(* IEC 61131-3 sources: SortJet_MasterSPS_Aufbau.fbsproj/09_Station/Stationen/_Allgemein, 5 files *)

(* ---- Arretierung_FB_V01_00_00.fb.st ---- *)
(* METADATA
{
	"v3Meta": {
		"objectGuid": "dcab1ddf-6c10-4772-a9bc-4c92780e70eb"
	}
}
*)
FUNCTION_BLOCK Arretierung_FB_V01_00_00
VAR_INPUT

  // EINGAENGE
  in_bStatusZylinderAusgefahren : BOOL;
  in_bStatusZylinderEingefahren : BOOL;

  // BOOLEAN
  bpReset                       : BOOL;
  bpAktivieren                  : BOOL;
  bpFreigabe                    : BOOL; // FREIGABE Pneumatik: ohne Freigabe Ventile aus, Bewegung pausiert (Startbefehl bleibt erhalten)
  bpStartAusfahren              : BOOL;
  bpStartEinfahren              : BOOL;

  // OPTIONEN
  bpAbfrageAusgefahrenVorhanden : BOOL := TRUE;   // Endlagensensor ausgefahren vorhanden, sonst gilt die Endlage nach tpBewegungszeit
  bpAbfrageEingefahrenVorhanden : BOOL := TRUE;   // Endlagensensor eingefahren vorhanden, sonst gilt die Endlage nach tpBewegungszeit
  tpBewegungszeit               : TIME := T#800MS; // Bewegungszeit je Richtung ohne Endlagensensor

END_VAR
VAR_OUTPUT
  // AUSGAENGE
  out_bZylinderAusfahren        : BOOL;
  out_bZylinderEinfahren        : BOOL;

  // BOOLEAN
  bpFehler                      : BOOL;
  bpDone                        : BOOL;

  // WORD
  wpFehlerNr                    : Fehlerkonstanten_EN;

  // ENUM
  epStatusZylinder : PneumatikZylinderStatus_EN;

END_VAR
VAR

  // STEPS
  steplAusfahren   : Steps_TE;
  steplEinfahren   : Steps_TE;

  // TIMER
  tonZylinderEingefahren     : TON; // EINSCHALTVERZOEGERUNG: Warten bis der Zylinder eingefahren wurde. Sonst wird ein Fehlerausgegeben
  tonZylinderAusgefahren     : TON; // EINSCHALTVERZOEGERUNG: Warten bis der Zylinder ausgefahren wurde. Sonst wird ein Fehlerausgegeben
  tonlBewegungszeitEinfahren : TON; // Bewegungszeit ohne Endlagensensor eingefahren
  tonlBewegungszeitAusfahren : TON; // Bewegungszeit ohne Endlagensensor ausgefahren

END_VAR

VAR CONSTANT

  // TIME
  cZEITLICHE_UEBERWACHUNG_BEWEGUNG_ZYLINDER : TIME := T#15s;

END_VAR
//-------------------------------------------------------------------------------------------------
// BAUSTEIN: RESET / DEAKTIVIERT
//-------------------------------------------------------------------------------------------------
(* Hinweis:
   - Reset oder deaktiviert: Ausgaenge aus, Ketten und Timer zuruecksetzen, Done und Fehler loeschen
   - Der Baustein setzt bpReset selbst zurueck, der Aufrufer wartet nicht auf Done
   - Ein deaktivierter Zylinder meldet kein Done; der Aufrufer verknuepft das Warten auf Done
     mit der Aktivierung aus der MK (z.B. Zylinder.bpDone OR NOT stStationsAufbau.bX)
*)
IF ( bpReset OR NOT bpAktivieren ) THEN

  out_bZylinderAusfahren := FALSE;
  out_bZylinderEinfahren := FALSE;

  bpStartAusfahren := FALSE;
  bpStartEinfahren := FALSE;

  steplAusfahren := STEP_0_E;
  steplEinfahren := STEP_0_E;

  tonZylinderAusgefahren( IN := FALSE );
  tonZylinderEingefahren( IN := FALSE );
  tonlBewegungszeitAusfahren( IN := FALSE );
  tonlBewegungszeitEinfahren( IN := FALSE );

  bpDone     := FALSE;
  bpFehler   := FALSE;
  wpFehlerNr := cMELDUNG_NULL;

  bpReset := FALSE;

  RETURN;

END_IF

//-------------------------------------------------------------------------------------------------
// BAUSTEIN: AKTIONEN
//-------------------------------------------------------------------------------------------------
(* Hinweis Freigabe Pneumatik:
   - Ohne Freigabe: Ventile aus, Ketten und Ueberwachungszeiten zuruecksetzen (kein Timeout-Fehler)
   - Der Startbefehl bleibt erhalten: kommt die Freigabe zurueck, wird die Bewegung neu gestartet
*)
IF NOT bpFreigabe THEN
  out_bZylinderAusfahren := FALSE;
  out_bZylinderEinfahren := FALSE;
  steplAusfahren := STEP_0_E;
  steplEinfahren := STEP_0_E;
  tonZylinderAusgefahren( IN := FALSE );
  tonZylinderEingefahren( IN := FALSE );
  tonlBewegungszeitAusfahren( IN := FALSE );
  tonlBewegungszeitEinfahren( IN := FALSE );
  bpDone := FALSE;
ELSE
  Ausfahren();
  Einfahren();
END_IF

//-------------------------------------------------------------------------------------------------
// STATUS DES ZYLINDERS
//-------------------------------------------------------------------------------------------------
(* Hinweis:
   - Status aus der Sensorik, soweit Endlagensensoren vorhanden sind
   - Ohne Sensor bleibt der Status, den die Schrittketten nach der Bewegungszeit setzen
*)
IF ( bpAbfrageAusgefahrenVorhanden AND bpAbfrageEingefahrenVorhanden ) THEN

  IF (      in_bStatusZylinderAusgefahren
       AND NOT in_bStatusZylinderEingefahren )
  THEN
    epStatusZylinder := eZylinderAusgefahren;
  ELSIF(    in_bStatusZylinderEingefahren
         AND NOT in_bStatusZylinderAusgefahren )
  THEN
    epStatusZylinder := eZylinderEingefahren;
  ELSE
    epStatusZylinder := eZylinderUndefiniert;
  END_IF

ELSIF ( bpAbfrageAusgefahrenVorhanden ) THEN

  IF ( in_bStatusZylinderAusgefahren ) THEN
    epStatusZylinder := eZylinderAusgefahren;
  ELSIF ( epStatusZylinder = eZylinderAusgefahren ) THEN
    epStatusZylinder := eZylinderUndefiniert;
  END_IF

ELSIF ( bpAbfrageEingefahrenVorhanden ) THEN

  IF ( in_bStatusZylinderEingefahren ) THEN
    epStatusZylinder := eZylinderEingefahren;
  ELSIF ( epStatusZylinder = eZylinderEingefahren ) THEN
    epStatusZylinder := eZylinderUndefiniert;
  END_IF

END_IF
END_FUNCTION_BLOCK

(* ---- Kippen_FB_V01_00_00.fb.st ---- *)
(* METADATA
{
	"v3Meta": {
		"objectGuid": "d572774f-9eb0-4642-b999-1d4bc3469776"
	}
}
*)
FUNCTION_BLOCK Kippen_FB_V01_00_00
VAR_INPUT

  // BOOLEAN *)
  bpAktivieren              : BOOL;
  bpFreigabe                : BOOL;
  bpReset                   : BOOL;
  bpReferenz                : BOOL;
  bpPositionieren           : BOOL;
  bpHandfahrenPlus          : BOOL;
  bpHandfahrenMinus         : BOOL;
  bpAutomatikAktiv          : BOOL;
  bpSensorEinlauf           : BOOL;
  bpSensorAuslauf           : BOOL;
  bpSensorEinlaufNachfolger : BOOL;
  bpSensorAuslaufVorgaenger : BOOL;
  bpTeilnehmerErreichbar    : BOOL;

  bpSensorNicht90Grad       : BOOL;

  bpLangsamKippen           : BOOL; // Umrichter: mit reduzierter Geschwindigkeit und Beschleunigung positionieren
  bpSensorNicht84Grad       : BOOL;

  // POINTER
  ppAntriebsInformationen : REFERENCE TO AntriebsInformationen;
  ppParameterBaustein     : REFERENCE TO Parameter_Kippen;

  // ENUM
  epZielPosition          : Kippen_EN; // Hinweis: Wird fuer die Absolut-Positionierung verwendet "bpStartAbsolutPositionierung"

  // STRUCT
  stStationsNummern       : Station_ST;

END_VAR
VAR_OUTPUT

  // BOOLEAN
  bpDone                       : BOOL;
  bpFehler                     : BOOL;
  bpInReferenz                 : BOOL;
  bpPositionierenAbgeschlossen : BOOL;

  // WORD
  wpFehlerNr                   : Fehlerkonstanten_EN; // FEHLER-AUSWERTUNG: Fehlernummer[Const] *)

  // ENUM *)
  epKippStatus                 : Kippen_EN; // Status: Gibt die aktuelle Position des Antriebs aus

END_VAR
VAR

  // BOOLEAN
  blErsterZyklus      : BOOL := TRUE;

  // REAL
  rlAntriebsZielPosition : REAL;

  // TIMER
  tonlFehlermeldungUnterdrueckenAntriebOK : TON;
  tonlMaxWarteZeit                        : TON;
  tonlMaxWarteAufResetErfolgreich         : TON;
  tonlAntriebNichtFreigegeben             : TON; // Ueberwachung: Antrieb nicht betriebsbereit
  tonlEndschalterFreifahren               : TON;
  tonlWarteSchrittEndschalterFreifahren   : TON;
  tofHardwareEndschalterFrei              : TOF;
  toflReglerFreigabeErhalten              : TOF;
  toflHardwareEndschalterFrei             : TOF;
  toflReset                               : TOF;

  // STEPS
  steplReset          : Steps_TE;
  steplReferenz       : Steps_TE;
  steplPositionieren  : Steps_TE;

  // Antrieb
  Antrieb : REFERENCE TO Rexroth_ctrlX_Drive_Eckelmann_MC_V01_02_02;

END_VAR

VAR
  // HARDWARE EINGÄNGE
  in_bMotorstarter_OK                 AT%I* : BOOL;
  in_bLS400V_OK                       AT%I* : BOOL;
  in_bLSBremse_OK                     AT%I* : BOOL;

  // HARDWARE AUSGÄNGE
  out_bKippen84Grad                   AT%Q* : BOOL;
  out_bKippen90Grad                   AT%Q* : BOOL;
  out_bBremseLoesen                   AT%Q* : BOOL;
  out_bReset                          AT%Q* : BOOL;

END_VAR

//-------------------------------------------------------------------------------------------------
// INITIALISIERUNG
//-------------------------------------------------------------------------------------------------
IF ( blErsterZyklus ) THEN

  IF ( __ISVALIDREF(ppAntriebsInformationen) ) THEN

    blErsterZyklus := FALSE;

    Antrieb REF= pgAntriebe[ppAntriebsInformationen.wAchsID];

    (* Hinweis:
       - Initialisierung Antriebsinformationen
    *)
    Antrieb.ppAntriebsInformationen REF= ppAntriebsInformationen;

    (* Hinweis:
       - Für die Zielpunktkontrolle muss im ersten Zyklus die Zielposition initialisiert werden
    *)
    Antrieb.rpZielPosition := Antrieb.rpIstPosition;

    (* Hinweis:
       - Antriebswerte vorinitialisieren
    *)
    Antrieb.rpGeschwindigkeit := ppAntriebsInformationen.rpMaxGeschwindigkeit;
    Antrieb.rpBeschleunigung  := ppAntriebsInformationen.rpMaxBeschleunigung;
    Antrieb.rpVerzoegerung    := ppAntriebsInformationen.rpMaxVerzoegerung;
    Antrieb.rpRuckzeit        := ppAntriebsInformationen.rpMaxRuckzeit;

  ELSE
    RETURN;
  END_IF

END_IF

//-------------------------------------------------------------------------------------------------
// DEAKTIVIEREN
//-------------------------------------------------------------------------------------------------
IF ( NOT bpAktivieren ) THEN

  bpDone                       := TRUE;
  bpInReferenz                 := TRUE;
  bpPositionierenAbgeschlossen := TRUE;

  epKippStatus := epZielPosition;

  bpFehler   := FALSE;
  wpFehlerNr := cMELDUNG_NULL;

  RETURN;

END_IF

//-------------------------------------------------------------------------------------------------
// BAUSTEIN: AKTIONEN
//-------------------------------------------------------------------------------------------------

(* Hinweis:
   - Kippbewegung
*)
IF (ppParameterBaustein.bKippenMitSchuetz ) THEN
  Kippen_Schuetz();
ELSE
  Positionieren();
END_IF

(* Hinweis:
   - Baisis- Aktionen
*)
Ausgaenge();
Meldungen();
Timer();
Reset();
Referenz();
Handbetrieb();

//-------------------------------------------------------------------------------------------------
// ZUWEISUNGEN UND BAUSTEINAUFRUFE
//-------------------------------------------------------------------------------------------------
// Antriebsfreigabe:
//    - Antrieb
toflReglerFreigabeErhalten( IN := (   bpPositionieren
                                    OR bpReferenz
                                    OR bpHandfahrenPlus
                                    OR bpHandfahrenMinus
                                    OR bpReset ),
                            PT := ppParameterBaustein.tZeitAntriebsfreigabeErhalten );

Antrieb.bpFreigabe        := ( bpFreigabe AND toflReglerFreigabeErhalten.Q );
IF ( NOT ( bpPositionieren AND bpLangsamKippen ) ) THEN
  Antrieb.rpRuckzeit      := ppAntriebsInformationen.rpMaxRuckzeit;
END_IF
Antrieb.stStationsNummern := stStationsNummern;
END_FUNCTION_BLOCK

(* ---- Messachse_FB_V01_00_00.fb.st ---- *)
(* METADATA
{
	"v3Meta": {
		"objectGuid": "ee8fce2f-1a3c-411c-afad-25d0a39b52dd"
	}
}
*)
FUNCTION_BLOCK Messachse_FB_V01_00_00
VAR_INPUT

  // BOOL
  bpAktivieren                             : BOOL;
  bpPositionierung                         : BOOL;
  bpVermessen_OberUndUnterkante_2_Sensoren : BOOL;
  bpVermessen_Oberkante_1_Sensor           : BOOL;
  bpReset                                  : BOOL;
  bpReferenz                               : BOOL;
  bpFreigabe                               : BOOL;
  bpHandfahrenPlus                         : BOOL;
  bpHandfahrenMinus                        : BOOL;
  bpBetriebsartHand                        : BOOL;
  bpFusstaster                             : BOOL;

 // REAL
  rpZielPosition                           : REAL;
  rpErwarteteScheibenHoehe                 : REAL;

  // STRUCT
  stStationsNummern                        : Station_ST;

  // POINTER
  ppAntriebsInformationen                  : REFERENCE TO AntriebsInformationen;
  ppParameterBaustein                      : REFERENCE TO Parameter_Messachse;

END_VAR
VAR_OUTPUT

  // BOOL
  bpDone                    : BOOL;
  bpFehler                  : BOOL;
  bpInReferenz              : BOOL;
  bprtScheibe               : BOOL;
  bpVermessenAbgeschlossen  : Bool;

  // WORD
  wpFehlerNr                : Fehlerkonstanten_EN;

  // REAL
  rpIstPosition             : REAL;
  rlScheibenunterkante      : REAL;
  rlScheibenoberkante       : REAL;
  rlMessErgebnis            : REAL;
  rlPositionAntriebBeiStart : REAL;
  rlBremsWeg                : REAL;

  // ENUM
  epGlashoehenTyp      : GlasHoehenTyp_EN;
  epGlashoehenTypMode2 : GlasHoehenTyp_EN;

END_VAR
VAR

  // BOOL
  blErsterZyklus                         : BOOL := TRUE;

  // REAL
  rlBremsPos                             : REAL;
  rlOffsetMinimumFrueherBremsen          : REAL := 150;
  rlOffsetMaximumFrueherBremsen          : REAL := 300;

  // TIMER
  tonlEndschalterFreifahren              : TON;
  tonlWarteSchrittEndschalterFreifahren  : TON;
  tonlMaxWarteAufResetErfolgreich        : TON;
  tonlAntriebNichtFreigegeben            : TON; // Ueberwachung: Antrieb nicht betriebsbereit
  tonlTimeoutUnterkante                  : TON;
  toflHardwareEndschalterFrei            : TOF;
  toflReglerFreigabeErhalten             : TOF;

  // STEPS
  steplPositionieren                     : Steps_TE;
  steplReferenz                          : Steps_TE;
  steplReset                             : Steps_TE;
  steplOberkante_1_Sensor                : Steps_TE;
  steplOberUndUnterkante_2_Sensoren      : Steps_TE;

  // Antrieb
  Antrieb : REFERENCE TO Rexroth_ctrlX_Drive_Eckelmann_MC_V01_02_02;

END_VAR

VAR_INPUT

  // HARDWARE EINGAENGE
  in_bSensorUnten                        : BOOL;
  in_bSensorOben                         : BOOL;
  in_bSensorUnterkante                   : BOOL;
  in_bEndschalterMin                     : BOOL; // Oeffner (TRUE = frei), gemappt; zum Umrichter ueber Signal-Steuerwort Bit 10, wirkt nur bei Endschalterquelle SPS

END_VAR
VAR CONSTANT

  // REAL
  cUEBERWACHUNG_WEGSTRECKE  : REAL := 40.0;

END_VAR

//-------------------------------------------------------------------------------------------------
// INITIALISIERUNG
//-------------------------------------------------------------------------------------------------
IF ( blErsterZyklus ) THEN

  IF ( __ISVALIDREF(ppAntriebsInformationen) ) THEN

    blErsterZyklus := FALSE;

    Antrieb REF= pgAntriebe[ppAntriebsInformationen.wAchsID];

    (* Hinweis:
       - Initialisierung Antriebsinformationen
    *)
    Antrieb.ppAntriebsInformationen REF= ppAntriebsInformationen;

    (* Hinweis:
       - Für die Zielpunktkontrolle muss im ersten Zyklus die Zielposition initialisiert werden
    *)
    Antrieb.rpZielPosition := Antrieb.rpIstPosition;

    (* Hinweis:
       - Antriebswerte vorinitialisieren
    *)
    Antrieb.rpGeschwindigkeit := ppAntriebsInformationen.rpMaxGeschwindigkeit;
    Antrieb.rpBeschleunigung  := ppAntriebsInformationen.rpMaxBeschleunigung;
    Antrieb.rpVerzoegerung    := ppAntriebsInformationen.rpMaxVerzoegerung;
    Antrieb.rpRuckzeit        := ppAntriebsInformationen.rpMaxRuckzeit;

  ELSE
    RETURN;
  END_IF

END_IF

//-------------------------------------------------------------------------------------------------
// DEAKTIVIEREN
//-------------------------------------------------------------------------------------------------
IF ( NOT bpAktivieren ) THEN

  bpDone := TRUE;

  (* Hinweis:
     - Ausnahmesituationen
  *)
  bpInReferenz := TRUE;
  bpFehler   := FALSE;
  wpFehlerNr := cMELDUNG_NULL;

  RETURN;

END_IF

//-------------------------------------------------------------------------------------------------
// IO's
//-------------------------------------------------------------------------------------------------
in_bSensorOben       := Antrieb.udipEingaengeUmrichter.cXG31_2_I_2;
in_bSensorUnten      := Antrieb.udipEingaengeUmrichter.cXG31_1_I_1;
in_bSensorUnterkante := Antrieb.udipEingaengeUmrichter.cXG37_4_I_6;
Antrieb.bpEndschalterMinExtern := in_bEndschalterMin;

//-------------------------------------------------------------------------------------------------
// BAUSTEIN: AKTIONEN
//-------------------------------------------------------------------------------------------------

Positionieren();
Vermessen_Oberkante_1_Sensor();
Vermessen_OberUndUnterkante_2_Sensoren();
Reset();
Referenz();
Handfunktion();

//-------------------------------------------------------------------------------------------------
// BAUSTEIN: AUSGAENGE
//-------------------------------------------------------------------------------------------------
// Ausgabe der Aktuellen Position
rpIstPosition := Antrieb.rpIstPosition;
bpInReferenz := Antrieb.bpIstReferenziert;

(* Hinweis:
   - Scheibenhoehe kontrollieren
*)
IF ( in_bSensorUnten AND NOT in_bSensorOben ) THEN
  epGlashoehenTyp := eGlasHoeheOK;

ELSE

  IF ( NOT in_bSensorUnten AND NOT in_bSensorOben ) THEN
    epGlashoehenTyp := eGlasZuNiedrig;

  ELSIF ( in_bSensorUnten AND  in_bSensorOben ) THEN
    epGlashoehenTyp := eGlasZuHoch;

  END_IF

END_IF

//-------------------------------------------------------------------------------------------------
// BAUSTEIN: AUFRUFE
//-------------------------------------------------------------------------------------------------
toflReglerFreigabeErhalten( IN := (   bpPositionierung
                                    OR bpReferenz
                                    OR bpHandfahrenPlus
                                    OR bpHandfahrenMinus
                                    OR bpVermessen_OberUndUnterkante_2_Sensoren
                                    OR bpVermessen_Oberkante_1_Sensor
                                    OR bpReset ),
                            PT := tgZeitAutoabschaltungEnergiesparModus );

Antrieb.bpFreigabe        := ( bpFreigabe AND toflReglerFreigabeErhalten.Q );
Antrieb.rpRuckzeit        := ppAntriebsInformationen.rpMaxRuckzeit;
Antrieb.stStationsNummern := stStationsNummern;

//-------------------------------------------------------------------------------------------------
// BAUSTEIN: AUSNAHMESITUATIONEN
//-------------------------------------------------------------------------------------------------
IF ( Antrieb.bpFehler
     AND NOT ( steplPositionieren = STEP_900_E
               OR steplOberUndUnterkante_2_Sensoren = STEP_900_E
               OR steplOberkante_1_Sensor = STEP_900_E
               OR steplReferenz    = STEP_900_E
               OR steplReset       = STEP_900_E ) )
THEN
  wpFehlerNR := cMELDUNG_ANTRIEB_MESSACHSE;
  bpFehler := TRUE;
END_IF
END_FUNCTION_BLOCK

(* ---- Querfahrt_FB_V01_00_00.fb.st ---- *)
(* METADATA
{
	"v3Meta": {
		"objectGuid": "62b3e7d5-59d7-4fa9-a26b-9f6c0e862cd9"
	}
}
*)
FUNCTION_BLOCK Querfahrt_FB_V01_00_00
VAR_INPUT

  // BOOLEAN
  bpAktivieren                           : BOOL;
  bpFreigabe                             : BOOL;
  bpAutomatikAktiv                       : BOOL;
  bpPositionieren                        : BOOL;
  bpReset                                : BOOL;
  bpReferenz                             : BOOL;
  bpHandfahrenPlus                       : BOOL;
  bpHandfahrenMinus                      : BOOL;

  bpSensorEinlauf                        : BOOL;
  bpSensorAuslauf                        : BOOL;
  bpSensorAuslaufVorgaenger              : BOOL;
  bpVerfahrfreigabe                      : BOOL := TRUE; // Externe Freigabe zum Verfahren (ohne Beschaltung TRUE)
  bpQuittungAuftragsstatusZurueckgesetzt : BOOL; // Auftrag wurde zurueckgesetzt
  bpReglungAktivSchalten                 : BOOL; // Da der Querfahrtantrieb keine Bremse hat, muss um die Position zu halten der Regler in Regelung stehen, sonst verschiebt sich die Station *)

  // REAL
  rpZielPosition                         : REAL;

  // POINTER
  ppParameterBaustein                    : REFERENCE TO Parameter_Querfahrt;
  ppAntriebsInformationen                : REFERENCE TO AntriebsInformationen;

  // STRUKTUR
  stStationsNummern                      : Station_ST;

END_VAR
VAR_OUTPUT

  // BOOLEAN
  bpDone                                 : BOOL;
  bpFehler                               : BOOL;
  bpAntrieblaeuft                        : BOOL;
  bpAuftragAktiv                         : BOOL;
  bpAuftragsstatusZuruecksetzen          : BOOL := FALSE;
  bpPositionierungGestartet              : BOOL := FALSE;
  bpPositionierungAbgeschlossen          : BOOL := FALSE;
  bpMinEndschalterBelegt                 : BOOL := FALSE;
  bpMaxEndschalterBelegt                 : BOOL := FALSE;
  bpZielPositionErreicht                 : BOOL;
  bpInReferenz                           : BOOL;

  // WORD
  wpFehlerNr                             : Fehlerkonstanten_EN;

  // REAL
  rpAktuellePosition                     : REAL;

END_VAR
VAR

  // BOOL
  blErsterZyklus                         : BOOL := TRUE;
  blVerfahrfreigabe                      : BOOL;
  blAbbruchPositionierung                : BOOL := FALSE;

  // STEPS
  steplPositionieren                     : Steps_TE;
  steplReferenz                          : Steps_TE;
  steplReset                             : Steps_TE;

  // TIMER
  tonlEndschalterFreifahren              : TON;
  tonlMaxWarteAufResetErfolgreich        : TON;
  toflHardwareEndschalterFrei            : TOF;
  toflReglerFreigabeErhalten             : TOF;

  // Antrieb
  Antrieb : REFERENCE TO Rexroth_ctrlX_Drive_Eckelmann_MC_V01_02_02;

END_VAR

//-------------------------------------------------------------------------------------------------
// INITIALISIERUNG
//-------------------------------------------------------------------------------------------------
IF ( blErsterZyklus ) THEN

  IF ( __ISVALIDREF(ppAntriebsInformationen) ) THEN

    blErsterZyklus := FALSE;

    Antrieb REF= pgAntriebe[ppAntriebsInformationen.wAchsID];

    (* Hinweis:
       - Initialisierung Antriebsinformationen
    *)
    Antrieb.ppAntriebsInformationen REF= ppAntriebsInformationen;

    (* Hinweis:
       - Für die Zielpunktkontrolle muss im ersten Zyklus die Zielposition initialisiert werden
    *)
    Antrieb.rpZielPosition := Antrieb.rpIstPosition;

    (* Hinweis:
       - Antriebswerte vorinitialisieren
    *)
    Antrieb.rpGeschwindigkeit := ppAntriebsInformationen.rpMaxGeschwindigkeit;
    Antrieb.rpBeschleunigung  := ppAntriebsInformationen.rpMaxBeschleunigung;
    Antrieb.rpVerzoegerung    := ppAntriebsInformationen.rpMaxVerzoegerung;
    Antrieb.rpRuckzeit        := ppAntriebsInformationen.rpMaxRuckzeit;

  ELSE
    RETURN;
  END_IF

END_IF

//-------------------------------------------------------------------------------------------------
// DEAKTIVIEREN
//-------------------------------------------------------------------------------------------------
IF ( NOT bpAktivieren ) THEN

  bpDone                        := TRUE;
  bpAuftragsstatusZuruecksetzen := FALSE;

  bpFehler   := FALSE;
  wpFehlerNr := cMELDUNG_NULL;

  RETURN;

END_IF

//-------------------------------------------------------------------------------------------------
// AKTIONEN
//-------------------------------------------------------------------------------------------------
// Verfahrfreigabe (lokal, der Eingang wird nicht ueberschrieben)
blVerfahrfreigabe :=     bpVerfahrfreigabe
                         AND NOT bpSensorEinlauf
                         AND NOT bpSensorAuslauf
                         AND NOT bpSensorAuslaufVorgaenger;

Verfahrlogik();
Positionieren();
Handfunktionen();
Reset();
Referenz();
Meldungen();

//-------------------------------------------------------------------------------------------------
// Freigabe zum Verfahren
//-------------------------------------------------------------------------------------------------
IF NOT blVerfahrfreigabe AND Antrieb.wpBetriebsart <> AntriebsBetriebsart_EN.RESET AND Antrieb.wpBetriebsart <> KEINE_FUNKTION THEN
  Antrieb.wpBetriebsart := KEINE_FUNKTION;
END_IF

//-------------------------------------------------------------------------------------------------
// Freigaben
//-------------------------------------------------------------------------------------------------
// Antriebsfreigabe
toflReglerFreigabeErhalten( IN := (   bpPositionieren
                                    OR bpReferenz
                                    OR bpHandfahrenPlus
                                    OR bpHandfahrenMinus
                                    OR bpReglungAktivSchalten // Da der Querfahrtantrieb keine Bremse hat, muss um die Position zu halten der Regler in Regelung stehen, sonst verschiebt sich die Station
                                    OR bpReset ),
                            PT := ppParameterBaustein.tZeitAntriebsfreigabeErhalten );

Antrieb.bpFreigabe        := ( bpFreigabe  AND toflReglerFreigabeErhalten.Q );
Antrieb.rpRuckzeit        := ppAntriebsInformationen.rpMaxRuckzeit;
Antrieb.stStationsNummern := stStationsNummern;

// Ausgänge
bpAuftragAktiv             := bpPositionieren;
rpAktuellePosition         := Antrieb.rpIstPosition;
bpAntrieblaeuft            := Antrieb.bpAntrieblaeuft;
bpInReferenz               := Antrieb.bpIstReferenziert;
bpMinEndschalterBelegt     := Antrieb.bpMinSchalterBelegt;
bpMaxEndschalterBelegt     := Antrieb.bpMaxSchalterBelegt;
bpPositionierungGestartet  := steplPositionieren > STEP_0_E;
bpPositionierungAbgeschlossen := bpDone AND NOT bpPositionieren;

// Positionsabfrage:
//    - Wurde die Zielposition aus dem Auftrag erreicht, bzw. stimmt die aktuelle Shuttleposition mit der
//      Position aus dem Auftrag ueberein.
bpZielPositionErreicht := ( ABS( rpZielposition - Antrieb.rpIstPosition ) <= rgMKZielPositionToleranz );
END_FUNCTION_BLOCK

(* ---- Scheibenmessung_FB_V01_00_00.fb.st ---- *)
(* METADATA
{
	"v3Meta": {
		"objectGuid": "c97c67c9-5e06-4086-aebd-8e091471f135"
	}
}
*)
FUNCTION_BLOCK Scheibenmessung_FB_V01_00_00
VAR_INPUT

  // BOOL
  bpReset                             : BOOL;
  bpGlasvermessung                    : BOOL;
  bpDrehrichtungsumkehrMessung        : BOOL; // FALSE = Positive Drehrichtung , TRUE = Negative Drehrichtung
  bpAuswahlSensorVorabScheibenmessung : BOOL;

  // REAL
  rpMessstrecke               : REAL;
  rpErwarteteScheibenLaenge   : REAL;
  rpFaktorBremswegverlaengern : REAL := 1.5;

  // POINTER
  ppAntrieb               : REFERENCE TO Rexroth_ctrlX_Drive_Eckelmann_MC_V01_02_02;
  pbpEinlaufSensor        : REFERENCE TO BOOL;
  pbpVorstopSensor        : REFERENCE TO BOOL;
  ppAntriebsInformationen : REFERENCE TO AntriebsInformationen;

  // ENUM
  epGlastyp               : GlasTyp_EN; // Default- oder Max-Scheibe, bestimmt die Ueberwachung des Einlaufsensors

  // STRUCT
  stStationsNummern       : Station_ST;

END_VAR
VAR_OUTPUT

  // BOOLEAN
  bpFehler                   : BOOL;
  bpGlasmessungAbgeschlossen : BOOL;

  // WORD
  wpFehlerNr                 : Fehlerkonstanten_EN;

  // REAL
  rpGemesseneGlaslaenge      : REAL;

END_VAR
VAR

  // REAL
  rlPositionAntriebBeiStart         : REAL;
  rlScheibenmessungErgebnis         : REAL;
  rlBremsWeg                        : REAL;
  rlMessergebnisMerker              : REAL;
  rlGefahrenerWeg                   : REAL;

  // STEPS
  steplGlasvermessung               : Steps_TE;

  // TIMER
  tonlAntriebNichtFreigegeben       : TON; // Ueberwachung: Antrieb nicht betriebsbereit

  // TRIGGER
  rtlMessung_OK                     : R_TRIG;

END_VAR

//-------------------------------------------------------------------------------------------------
// BAUSTEIN: SCHEIBENMESSUNG (LAENGE)
//-------------------------------------------------------------------------------------------------
(* Hinweis:
   - Reset setzt alles zurueck
*)
IF ( bpReset ) THEN
  bpGlasvermessung := FALSE;
  bpReset          := FALSE;

  wpFehlerNr := cMELDUNG_NULL;
  bpFehler   := FALSE;

  bpGlasmessungAbgeschlossen := FALSE;

ELSE
  Messung();

END_IF
END_FUNCTION_BLOCK
